(* Tx/Rx (string data) fifo control function block *)
FUNCTION_BLOCK FB_UDPFrameFIFO
VAR_INPUT
	bLog		: BOOL := FALSE;(* TRUE => Enable log message output, FALSE => Disable *)
	sPrefix		: STRING := 'Unknown::';(* Log message description string (allows the identification of log message source) *)
	stPut		: ST_UDPFrameEntry;(* Frame entry to add (write) to the buffer *)
END_VAR
VAR_OUTPUT
	bOk			: BOOL;(* TRUE = New entry added or removed succesfully, FALSE = Fifo overflow or fifo empty *)
	stGet		: ST_UDPFrameEntry;(* Frame entry removed (read) from fifo *)
	nCount		: UDINT := 0;(* Number of fifo entries *)
END_VAR
VAR
	fbBuffer 	: FB_MemRingBuffer;(* Basic (lower level) string buffer control function block *)
	buffer		: ARRAY[0..UDP_RX_BUFFER_SIZE] OF BYTE;(* Internal buffer memory *)
	fbCriticalSection:	FB_IecCriticalSection; (* Critical Section required for thread-safety *)
END_VAR

ACTION AddTail:
(* Adds new fifo entry *)
// IF fbCriticalSection.Enter() THEN
	fbBuffer.A_AddTail( pBuffer:= ADR(buffer), cbBuffer:= SIZEOF(buffer),
					pWrite:= ADR( stPut ), cbWrite := SIZEOF( stPut ), 
					bOk=>bOk, nCount=>nCount );
					
// 	fbCriticalSection.Leave();
// END_IF
// IF bOk AND bLog THEN(* Log message *)
// 	ADSLOGSTR( ADSLOG_MSGTYPE_HINT OR ADSLOG_MSGTYPE_LOG, 
// 			CONCAT( CONCAT( sPrefix, SOCKETADDR_TO_STRING(stPut.stRemoteAddr) ), '>>"%s"' ),
// 			stPut.sMessage );
// END_IF
END_ACTION

ACTION Clear:
(* Clears all fifo entries *)
// stGet.sMessage := 0;
// IF fbCriticalSection.Enter() THEN
	MEMSET(ADR(stGet.sMessage), 0, SIZEOF(stGet.sMessage));
	stGet.stRemoteAddr.nPort := 0;
	stGet.stRemoteAddr.sAddr := '';
	fbBuffer.A_Reset( pBuffer := ADR( buffer ), cbBuffer := SIZEOF( buffer ), bOk=>bOk, nCount=>nCount ); 
	
// 	fbCriticalSection.Leave();
// END_IF
END_ACTION

ACTION RemoveHead:
(* Removes oldest fifo entry *)

// IF fbCriticalSection.Enter() THEN
	IF nCount = 0 THEN
		MEMSET(ADR(stGet.sMessage), 0, SIZEOF(stGet.sMessage));
		stGet.stRemoteAddr.nPort := 0;
		stGet.stRemoteAddr.sAddr := '';
		bOk := FALSE;
		RETURN;
	END_IF
	
	fbBuffer.A_RemoveHead( pBuffer:= ADR(buffer), cbBuffer:= SIZEOF(buffer),
							pRead := ADR( stGet ), cbRead := SIZEOF( stGet ),
							bOk=>bOk, nCount=>nCount );
// 	fbCriticalSection.Leave();
// END_IF
END_ACTION

METHOD TEMPRemoveHead : BOOL
VAR_IN_OUT
	stGet	: ST_UDPFrameEntry;
END_VAR
VAR_INPUT
END_VAR
VAR_OUTPUT
	bOk		: BOOL;
END_VAR
IF fbCriticalSection.Enter() THEN
	IF nCount = 0 THEN
		MEMSET(ADR(stGet.sMessage), 0, SIZEOF(stGet.sMessage));
		stGet.stRemoteAddr.nPort := 0;
		stGet.stRemoteAddr.sAddr := '';
		bOk := FALSE;
		RETURN;
	END_IF
	
	fbBuffer.A_RemoveHead( pBuffer:= ADR(buffer), cbBuffer:= SIZEOF(buffer),
							pRead := ADR( stGet ), cbRead := SIZEOF( stGet ),
							bOk=>bOk, nCount=>nCount );
	fbCriticalSection.Leave();
END_IF
END_METHOD

END_FUNCTION_BLOCK

(* stored: Version 1.1.0.1
   POU FB_UDPFrameFIFO: Id {bdee9b83-07c8-47a7-8ab0-131de1831bda}, SpecialFunc None
   Action AddTail: Id {46e5920e-6c9c-4fa8-ba62-0a0a847d37eb}
   Action Clear: Id {665a0510-09d5-4318-8a19-fd1f2b292181}
   Action RemoveHead: Id {13ea9795-e95e-4f4f-a519-2dbc2dda7a42}
   Method TEMPRemoveHead: Id {b657f026-5eb2-4f4a-b09f-8934a623ef4e} *)
